(* IEC 61131-3 sources: plcassist-cli/packages/volt-lsp-iec/test-corpus/awa-palletizer/Device/Plc Logic/Application/Library Manager/ElementCollections, 110 files *)

(* ---- CONSTANTS.gvl ---- *)
VAR_GLOBAL
	GC_TREENODEFACTORY : TreeNodeFactory := STRUCT();
	GC_LINKEDOBJECTREFERENCEFACTORY : LinkedObjectReferenceFactory := STRUCT();
END_VAR

(* ---- VARIABLES.gvl ---- *)
VAR_GLOBAL
	G_LOCKWAITTIME : SYSTIME := 300;
	G_NULLELEMENT : NullElement;
END_VAR

(* ---- IBOOLELEMENT.itf ---- *)
INTERFACE IBOOLELEMENT
END_INTERFACE

(* ---- ICOLLECTION.itf ---- *)
INTERFACE ICOLLECTION
END_INTERFACE

METHOD ADDELEMENT : COLLECTION_ERROR
VAR_INPUT
	ITFELEMENT : IElement;
END_VAR
END_METHOD

METHOD CONTAINSELEMENT : COLLECTION_ERROR
VAR_INPUT
	ITFELEMENT : IElement;
END_VAR
VAR_OUTPUT
	XRESULT : BOOL;
END_VAR
END_METHOD

METHOD COUNTELEMENTS : UDINT
END_METHOD

METHOD ELEMENTITERATOR : COLLECTION_ERROR
VAR_INPUT
	ITFITERATOR : IIterator;
END_VAR
END_METHOD

METHOD REMOVEALLELEMENTS : COLLECTION_ERROR
END_METHOD

METHOD REMOVEELEMENT : COLLECTION_ERROR
VAR_INPUT
	ITFELEMENT : IElement;
END_VAR
END_METHOD

(* ---- ICONTAINSVALUE.itf ---- *)
INTERFACE ICONTAINSVALUE
END_INTERFACE

METHOD CONTAINSVALUE : COLLECTION_ERROR
VAR_INPUT
	ITFELEMENT : IElement;
END_VAR
VAR_OUTPUT
	XRESULT : BOOL;
END_VAR
END_METHOD

(* ---- IDINTELEMENT.itf ---- *)
INTERFACE IDINTELEMENT
END_INTERFACE

(* ---- IDOUBLELINKEDLIST.itf ---- *)
INTERFACE IDOUBLELINKEDLIST
END_INTERFACE

METHOD REMOVEFIRSTELEMENT : COLLECTION_ERROR
END_METHOD

METHOD REMOVELASTELEMENT : COLLECTION_ERROR
END_METHOD

(* ---- IDOUBLELINKEDLIST2.itf ---- *)
INTERFACE IDOUBLELINKEDLIST2
END_INTERFACE

METHOD SAFEELEMENTITERATOR : COLLECTION_ERROR
VAR_INPUT
	ITFITERATOR : ISafeLinkedListIterator;
END_VAR
END_METHOD

(* ---- IELEMENT.itf ---- *)
INTERFACE IELEMENT
END_INTERFACE

METHOD ELEMENTCOMPARETO : INT
VAR_INPUT
	ITFELEMENT : IElement;
END_VAR
END_METHOD

METHOD ELEMENTEQUALS : BOOL
VAR_INPUT
	ITFELEMENT : IElement;
END_VAR
END_METHOD

METHOD ELEMENTHASHCODE : LINT
END_METHOD

(* ---- IINTELEMENT.itf ---- *)
INTERFACE IINTELEMENT
END_INTERFACE

(* ---- IITERATOR.itf ---- *)
INTERFACE IITERATOR
END_INTERFACE

METHOD HASNEXT : BOOL
END_METHOD

METHOD NEXT : COLLECTION_ERROR
VAR_OUTPUT
	ITFELEMENT : IElement;
END_VAR
END_METHOD

(* ---- ILINKEDLISTITERATOR.itf ---- *)
INTERFACE ILINKEDLISTITERATOR
END_INTERFACE

(* ---- ILINKEDOBJECTREFERENCE.itf ---- *)
INTERFACE ILINKEDOBJECTREFERENCE
END_INTERFACE

(* ---- ILINTELEMENT.itf ---- *)
INTERFACE ILINTELEMENT
END_INTERFACE

(* ---- ILIST.itf ---- *)
INTERFACE ILIST
END_INTERFACE

METHOD GETELEMENTAT : COLLECTION_ERROR
VAR_INPUT
	UDIPOSITION : UDINT;
END_VAR
VAR_OUTPUT
	ITFELEMENT : IElement;
END_VAR
END_METHOD

METHOD GETELEMENTPOSITION : COLLECTION_ERROR
VAR_INPUT
	ITFELEMENT : IElement;
END_VAR
VAR_OUTPUT
	UDIPOSITION : UDINT;
END_VAR
END_METHOD

METHOD INSERTELEMENTAT : COLLECTION_ERROR
VAR_INPUT
	UDIPOSITION : UDINT;
	ITFELEMENT : IElement;
END_VAR
END_METHOD

METHOD REMOVEELEMENTAT : COLLECTION_ERROR
VAR_INPUT
	UDIPOSITION : UDINT;
END_VAR
END_METHOD

METHOD SETELEMENTAT : COLLECTION_ERROR
VAR_INPUT
	UDIPOSITION : UDINT;
	ITFELEMENT : IElement;
END_VAR
END_METHOD

(* ---- ILIST2.itf ---- *)
INTERFACE ILIST2
END_INTERFACE

(* ---- ILIST3.itf ---- *)
INTERFACE ILIST3
END_INTERFACE

METHOD SAFEELEMENTITERATOR : COLLECTION_ERROR
VAR_INPUT
	ITFITERATOR : ISafeListIterator;
END_VAR
END_METHOD

(* ---- ILISTITERATOR.itf ---- *)
INTERFACE ILISTITERATOR
END_INTERFACE

(* ---- ILOCKABLE.itf ---- *)
INTERFACE ILOCKABLE
END_INTERFACE

METHOD LOCK : BOOL
END_METHOD

METHOD RELEASELOCK
END_METHOD

(* ---- IMAP.itf ---- *)
INTERFACE IMAP
END_INTERFACE

METHOD ADDKEYVALUEPAIR : COLLECTION_ERROR
VAR_INPUT
	ITFKEY : IElement;
	ITFVALUE : IElement;
END_VAR
END_METHOD

METHOD CONTAINSKEY : COLLECTION_ERROR
VAR_INPUT
	ITFKEY : IElement;
END_VAR
VAR_OUTPUT
	XRESULT : BOOL;
END_VAR
END_METHOD

METHOD COUNTKEYS : UDINT
END_METHOD

METHOD GETELEMENTBYKEY : COLLECTION_ERROR
VAR_INPUT
	ITFKEY : IElement;
END_VAR
VAR_OUTPUT
	ITFVALUE : IElement;
END_VAR
END_METHOD

METHOD KEYS : COLLECTION_ERROR
VAR_INPUT
	ITFITERATOR : IIterator;
END_VAR
END_METHOD

METHOD REMOVEBYKEY : COLLECTION_ERROR
VAR_INPUT
	ITFKEY : IElement;
END_VAR
END_METHOD

METHOD VALUES : COLLECTION_ERROR
VAR_INPUT
	ITFITERATOR : IIterator;
END_VAR
END_METHOD

(* ---- IMAP2.itf ---- *)
INTERFACE IMAP2
END_INTERFACE

METHOD REMOVEALLELEMENTS : COLLECTION_ERROR
END_METHOD

(* ---- IMAP3.itf ---- *)
INTERFACE IMAP3
END_INTERFACE

METHOD SAFEKEYS : COLLECTION_ERROR
VAR_INPUT
	ITFITERATOR : ISafeListIterator;
END_VAR
END_METHOD

METHOD SAFEVALUES : COLLECTION_ERROR
VAR_INPUT
	ITFITERATOR : ISafeListIterator;
END_VAR
END_METHOD

(* ---- IMODCOUNTER.itf ---- *)
INTERFACE IMODCOUNTER
END_INTERFACE

(* ---- INULLELEMENT.itf ---- *)
INTERFACE INULLELEMENT
END_INTERFACE

(* ---- IOBJECTREFERENCE.itf ---- *)
INTERFACE IOBJECTREFERENCE
END_INTERFACE

(* ---- IONLINECHANGESAFELINKEDLISTELEMENT.itf ---- *)
INTERFACE IONLINECHANGESAFELINKEDLISTELEMENT
END_INTERFACE

METHOD UPDATEELEMENT
VAR_INPUT
	ITFELEMENT : IElement;
END_VAR
END_METHOD

(* ---- IQUEUE.itf ---- *)
INTERFACE IQUEUE
END_INTERFACE

METHOD PEEK : COLLECTION_ERROR
VAR_OUTPUT
	ITFELEMENT : IElement;
END_VAR
END_METHOD

METHOD POLL : COLLECTION_ERROR
VAR_OUTPUT
	ITFELEMENT : IElement;
END_VAR
END_METHOD

(* ---- IQUEUE2.itf ---- *)
INTERFACE IQUEUE2
END_INTERFACE

(* ---- IQUEUE3.itf ---- *)
INTERFACE IQUEUE3
END_INTERFACE

METHOD SAFEELEMENTITERATOR : COLLECTION_ERROR
VAR_INPUT
	ITFITERATOR : ISafeListIterator;
END_VAR
END_METHOD

(* ---- ISAFEITERATOR.itf ---- *)
INTERFACE ISAFEITERATOR
END_INTERFACE

METHOD NEXT : COLLECTION_ERROR
VAR_OUTPUT
	ITFELEMENT : IElement;
END_VAR
END_METHOD

(* ---- ISAFELINKEDLISTITERATOR.itf ---- *)
INTERFACE ISAFELINKEDLISTITERATOR
END_INTERFACE

(* ---- ISAFELISTITERATOR.itf ---- *)
INTERFACE ISAFELISTITERATOR
END_INTERFACE

(* ---- ISORTEDLIST.itf ---- *)
INTERFACE ISORTEDLIST
END_INTERFACE

METHOD ADDELEMENTWITHOUTSORTING : COLLECTION_ERROR
VAR_INPUT
	ITFELEMENT : IElement;
END_VAR
END_METHOD

METHOD SORT : COLLECTION_ERROR
END_METHOD

(* ---- ISORTEDLIST2.itf ---- *)
INTERFACE ISORTEDLIST2
END_INTERFACE

(* ---- ISORTEDLIST3.itf ---- *)
INTERFACE ISORTEDLIST3
END_INTERFACE

METHOD SAFEELEMENTITERATOR : COLLECTION_ERROR
VAR_INPUT
	ITFITERATOR : ISafeListIterator;
END_VAR
END_METHOD

(* ---- ISTACK.itf ---- *)
INTERFACE ISTACK
END_INTERFACE

METHOD PEEK : COLLECTION_ERROR
VAR_OUTPUT
	ITFELEMENT : IElement;
END_VAR
END_METHOD

METHOD POP : COLLECTION_ERROR
VAR_OUTPUT
	ITFELEMENT : IElement;
END_VAR
END_METHOD

(* ---- ISTACK2.itf ---- *)
INTERFACE ISTACK2
END_INTERFACE

(* ---- ISTACK3.itf ---- *)
INTERFACE ISTACK3
END_INTERFACE

METHOD SAFEELEMENTITERATOR : COLLECTION_ERROR
VAR_INPUT
	ITFITERATOR : ISafeListIterator;
END_VAR
END_METHOD

(* ---- ISTRINGELEMENT.itf ---- *)
INTERFACE ISTRINGELEMENT
END_INTERFACE

(* ---- ITIMEELEMENT.itf ---- *)
INTERFACE ITIMEELEMENT
END_INTERFACE

(* ---- ITREENODE.itf ---- *)
INTERFACE ITREENODE
END_INTERFACE

METHOD ADDCHILD : COLLECTION_ERROR
VAR_INPUT
	ITFELEMENT : IElement;
END_VAR
VAR_OUTPUT
	ITFTREENODE : ITreeNode;
END_VAR
END_METHOD

METHOD CHILDREN : COLLECTION_ERROR
VAR_INPUT
	ITFITERATOR : IIterator;
END_VAR
END_METHOD

METHOD CONTAINSCHILD : COLLECTION_ERROR
VAR_INPUT
	ITFELEMENT : IElement;
END_VAR
VAR_OUTPUT
	XRESULT : BOOL;
END_VAR
END_METHOD

METHOD COUNTCHILDREN : UDINT
END_METHOD

METHOD MOVENODE : COLLECTION_ERROR
VAR_INPUT
	ITFTARGETTREENODE : ITreeNode;
END_VAR
END_METHOD

METHOD PARENT : COLLECTION_ERROR
VAR_OUTPUT
	ITFPARENT : ITreeNode;
END_VAR
END_METHOD

METHOD REMOVECHILD : COLLECTION_ERROR
VAR_INPUT
	ITFELEMENT : IElement;
END_VAR
END_METHOD

METHOD ROOTNODE : COLLECTION_ERROR
VAR_OUTPUT
	ITFROOTNODE : ITreeNode;
END_VAR
END_METHOD

(* ---- ITREENODE2.itf ---- *)
INTERFACE ITREENODE2
END_INTERFACE

METHOD SAFECHILDREN : COLLECTION_ERROR
VAR_INPUT
	ITFITERATOR : ISafeLinkedListIterator;
END_VAR
END_METHOD

(* ---- IUDINTELEMENT.itf ---- *)
INTERFACE IUDINTELEMENT
END_INTERFACE

(* ---- IUINTELEMENT.itf ---- *)
INTERFACE IUINTELEMENT
END_INTERFACE

(* ---- IULINTELEMENT.itf ---- *)
INTERFACE IULINTELEMENT
END_INTERFACE

(* ---- IWSTRINGELEMENT.itf ---- *)
INTERFACE IWSTRINGELEMENT
END_INTERFACE

(* ---- COMPARESTRING.fun ---- *)
FUNCTION COMPARESTRING : INT
VAR_INPUT
	PS1 : POINTER TO STRING;
	PS2 : POINTER TO STRING;
END_VAR
END_FUNCTION

(* ---- COMPAREWSTRING.fun ---- *)
FUNCTION COMPAREWSTRING : INT
VAR_INPUT
	PW1 : POINTER TO WSTRING;
	PW2 : POINTER TO WSTRING;
END_VAR
END_FUNCTION

(* ---- GETLIBVERSION.fun ---- *)
FUNCTION GETLIBVERSION : VERSION
END_FUNCTION

(* ---- GETLIBVERSIONNUMBER.fun ---- *)
FUNCTION GETLIBVERSIONNUMBER : DWORD
END_FUNCTION

(* ---- HASHCODEFROMSTRING.fun ---- *)
FUNCTION HASHCODEFROMSTRING : UDINT
VAR_INPUT
	PSIN : POINTER TO STRING;
END_VAR
END_FUNCTION

(* ---- HASHCODEFROMWSTRING.fun ---- *)
FUNCTION HASHCODEFROMWSTRING : UDINT
VAR_INPUT
	PWIN : POINTER TO WSTRING;
END_VAR
END_FUNCTION

(* ---- ISLIBRELEASED.fun ---- *)
FUNCTION ISLIBRELEASED : BOOL
END_FUNCTION

(* ---- BOOLDATA.fb ---- *)
FUNCTION_BLOCK BOOLDATA EXTENDS InstanceData
VAR_INPUT
	XVALUE : BOOL;
END_VAR
END_FUNCTION_BLOCK

(* ---- BOOLELEMENT.fb ---- *)
FUNCTION_BLOCK BOOLELEMENT EXTENDS InstanceBase
VAR_INPUT
	XVALUE : BOOL;
END_VAR
VAR
	BOOLVALUE : BOOL;
END_VAR
END_FUNCTION_BLOCK

METHOD ELEMENTCOMPARETO : INT
VAR_INPUT
	ITFELEMENT : IElement;
END_VAR
END_METHOD

METHOD ELEMENTEQUALS : BOOL
VAR_INPUT
	ITFELEMENT : IElement;
END_VAR
END_METHOD

METHOD ELEMENTHASHCODE : LINT
END_METHOD

METHOD PRVINSTINIT : FBF.ERROR
VAR_INPUT
	ITFDATA : FBF.IData;
END_VAR
END_METHOD

(* ---- BOOLELEMENTFACTORY.fb ---- *)
FUNCTION_BLOCK BOOLELEMENTFACTORY EXTENDS FactoryBase
VAR
	PRVINSTCOUNT : CAA.COUNT;
	PRVINSTPOOLEXTENDSFACTOR : USINT;
	PRVINSTSIZE : CAA.SIZE;
END_VAR
END_FUNCTION_BLOCK

METHOD CREATE : IBoolElement
VAR_INPUT
	XVALUE : BOOL;
END_VAR
VAR_OUTPUT
	EERROR : FBF.ERROR;
END_VAR
END_METHOD

(* ---- DINTDATA.fb ---- *)
FUNCTION_BLOCK DINTDATA EXTENDS InstanceData
VAR_INPUT
	DIVALUE : DINT;
END_VAR
END_FUNCTION_BLOCK

(* ---- DINTELEMENT.fb ---- *)
FUNCTION_BLOCK DINTELEMENT EXTENDS InstanceBase
VAR_INPUT
	DIVALUE : DINT;
END_VAR
VAR
	DINTVALUE : DINT;
END_VAR
END_FUNCTION_BLOCK

METHOD ELEMENTCOMPARETO : INT
VAR_INPUT
	ITFELEMENT : IElement;
END_VAR
END_METHOD

METHOD ELEMENTEQUALS : BOOL
VAR_INPUT
	ITFELEMENT : IElement;
END_VAR
END_METHOD

METHOD ELEMENTHASHCODE : LINT
END_METHOD

METHOD PRVINSTINIT : FBF.ERROR
VAR_INPUT
	ITFDATA : FBF.IData;
END_VAR
END_METHOD

(* ---- DINTELEMENTFACTORY.fb ---- *)
FUNCTION_BLOCK DINTELEMENTFACTORY EXTENDS FactoryBase
VAR
	PRVINSTCOUNT : CAA.COUNT;
	PRVINSTPOOLEXTENDSFACTOR : USINT;
	PRVINSTSIZE : CAA.SIZE;
END_VAR
END_FUNCTION_BLOCK

METHOD CREATE : IDintElement
VAR_INPUT
	DIVALUE : DINT;
END_VAR
VAR_OUTPUT
	EERROR : FBF.ERROR;
END_VAR
END_METHOD

(* ---- HASHTABLE.fb ---- *)
FUNCTION_BLOCK HASHTABLE EXTENDS InstanceBase
VAR_INPUT
	PAELEMENTS : POINTER TO KeyValuePair;
	PALINKEDELEMENTS : POINTER TO KeyValuePair;
	PAITERATORELEMENTS : POINTER TO IElement;
	UDIMAXELEMENTS : UDINT;
END_VAR
VAR
	_UDICOUNT : UDINT;
	_XWPOINTERTOTHIS : __XWORD := THIS;
	_BYLOCK : BYTE;
	_ULINTCOUNTMODS : ULINT;
	_UIGROWFACTOR : UINT := 1;
	_UIPREALLOCATION : UINT := 100;
	_LOCKWAITTIME : SYSTIME := Variables.g_LockWaitTime;
	COUNTMODIFICATIONS : ULINT;
	LOCKWAITTIME : SYSTIME;
END_VAR
END_FUNCTION_BLOCK

METHOD ADDKEYVALUEPAIR : COLLECTION_ERROR
VAR_INPUT
	ITFKEY : IElement;
	ITFVALUE : IElement;
END_VAR
END_METHOD

METHOD ADDKEYVALUEPAIRINTERNAL : COLLECTION_ERROR
VAR_INPUT
	ITFKEY : IElement;
	ITFVALUE : IElement;
	XINCREF : BOOL;
END_VAR
END_METHOD

METHOD CONTAINSKEY : COLLECTION_ERROR
VAR_INPUT
	ITFKEY : IElement;
END_VAR
VAR_OUTPUT
	XRESULT : BOOL;
END_VAR
END_METHOD

METHOD CONTAINSKEYINTERNAL : COLLECTION_ERROR
VAR_INPUT
	ITFKEY : IElement;
END_VAR
VAR_OUTPUT
	XRESULT : BOOL;
END_VAR
END_METHOD

METHOD COUNTKEYS : UDINT
END_METHOD

METHOD DISPOSE : BOOL
END_METHOD

METHOD ELEMENTCOMPARETO : INT
VAR_INPUT
	ITFELEMENT : IElement;
END_VAR
END_METHOD

METHOD ELEMENTEQUALS : BOOL
VAR_INPUT
	ITFELEMENT : IElement;
END_VAR
END_METHOD

METHOD ELEMENTHASHCODE : LINT
END_METHOD

METHOD GETARRAYINDEX : UDINT
VAR_INPUT
	ITFKEY : IElement;
END_VAR
END_METHOD

METHOD GETELEMENTBYKEY : COLLECTION_ERROR
VAR_INPUT
	ITFKEY : IElement;
END_VAR
VAR_OUTPUT
	ITFVALUE : IElement;
END_VAR
END_METHOD

METHOD KEYS : COLLECTION_ERROR
VAR_INPUT
	ITFITERATOR : IIterator;
END_VAR
END_METHOD

METHOD LOCK : BOOL
END_METHOD

METHOD NEXTFREELINKEDELEMENT : COLLECTION_ERROR
VAR_OUTPUT
	PKEYVALUEPAIR : POINTER TO KeyValuePair;
END_VAR
END_METHOD

METHOD REALLOC : BOOL
END_METHOD

METHOD RELEASELOCK
END_METHOD

METHOD REMOVEALLELEMENTS : COLLECTION_ERROR
END_METHOD

METHOD REMOVEBYKEY : COLLECTION_ERROR
VAR_INPUT
	ITFKEY : IElement;
END_VAR
END_METHOD

METHOD SAFEKEYS : COLLECTION_ERROR
VAR_INPUT
	ITFITERATOR : ISafeListIterator;
END_VAR
END_METHOD

METHOD SAFEVALUES : COLLECTION_ERROR
VAR_INPUT
	ITFITERATOR : ISafeListIterator;
END_VAR
END_METHOD

METHOD VALUES : COLLECTION_ERROR
VAR_INPUT
	ITFITERATOR : IIterator;
END_VAR
END_METHOD

METHOD PRVINSTINIT : FBF.ERROR
VAR_INPUT
	ITFDATA : FBF.IData;
END_VAR
END_METHOD

(* ---- HASHTABLEARGS.fb ---- *)
FUNCTION_BLOCK HASHTABLEARGS EXTENDS InstanceData
VAR_INPUT
	PAELEMENTS : POINTER TO KeyValuePair;
	PALINKEDELEMENTS : POINTER TO KeyValuePair;
	PAITERATORELEMENTS : POINTER TO IElement;
	UDIMAXELEMENTS : UDINT;
	UIGROWFACTOR : UINT;
	UIPREALLOCATION : UINT;
END_VAR
END_FUNCTION_BLOCK

(* ---- HASHTABLEFACTORY.fb ---- *)
FUNCTION_BLOCK HASHTABLEFACTORY EXTENDS FactoryBase
VAR
	PRVINSTCOUNT : CAA.COUNT;
	PRVINSTPOOLEXTENDSFACTOR : USINT;
	PRVINSTSIZE : CAA.SIZE;
END_VAR
END_FUNCTION_BLOCK

METHOD CREATE : IMap3
VAR_INPUT
	UDIMAXELEMENTS : UDINT;
END_VAR
VAR_OUTPUT
	EERROR : FBF.ERROR;
END_VAR
END_METHOD

METHOD CREATEDYNAMICHASHTABLE : IMap2
VAR_INPUT
	UDIINITIALSIZE : UDINT;
	UIGROWFACTOR : UINT;
END_VAR
VAR_OUTPUT
	EERROR : FBF.ERROR;
END_VAR
END_METHOD

METHOD CREATEDYNAMICHASHTABLEPREALLOC : IMap2
VAR_INPUT
	UDIINITIALSIZE : UDINT;
	UIGROWFACTOR : UINT;
	UIPREALLOCATION : UINT;
END_VAR
VAR_OUTPUT
	EERROR : FBF.ERROR;
END_VAR
END_METHOD

(* ---- INTDATA.fb ---- *)
FUNCTION_BLOCK INTDATA EXTENDS InstanceData
VAR_INPUT
	IVALUE : INT;
END_VAR
END_FUNCTION_BLOCK

(* ---- INTELEMENT.fb ---- *)
FUNCTION_BLOCK INTELEMENT EXTENDS InstanceBase
VAR_INPUT
	IVALUE : INT;
END_VAR
VAR
	INTVALUE : INT;
END_VAR
END_FUNCTION_BLOCK

METHOD ELEMENTCOMPARETO : INT
VAR_INPUT
	ITFELEMENT : IElement;
END_VAR
END_METHOD

METHOD ELEMENTEQUALS : BOOL
VAR_INPUT
	ITFELEMENT : IElement;
END_VAR
END_METHOD

METHOD ELEMENTHASHCODE : LINT
END_METHOD

METHOD PRVINSTINIT : FBF.ERROR
VAR_INPUT
	ITFDATA : FBF.IData;
END_VAR
END_METHOD

(* ---- INTELEMENTFACTORY.fb ---- *)
FUNCTION_BLOCK INTELEMENTFACTORY EXTENDS FactoryBase
VAR
	PRVINSTCOUNT : CAA.COUNT;
	PRVINSTPOOLEXTENDSFACTOR : USINT;
	PRVINSTSIZE : CAA.SIZE;
END_VAR
END_FUNCTION_BLOCK

METHOD CREATE : IIntElement
VAR_INPUT
	IVALUE : INT;
END_VAR
VAR_OUTPUT
	EERROR : FBF.ERROR;
END_VAR
END_METHOD

(* ---- LINKEDLIST.fb ---- *)
FUNCTION_BLOCK LINKEDLIST EXTENDS InstanceBase
VAR
	_SNAME : STRING := 'LinkedList';
	_RESULT : RTS_IEC_RESULT;
	_XWPOINTERTOTHIS : __XWORD := THIS;
	_BYLOCK : BYTE;
	_ULINTCOUNTMODS : ULINT;
	_ITFFIRSTLINKEDOBJECTREFERENCE : ILinkedObjectReference := 0;
	_ITFLASTLINKEDOBJECTREFERENCE : ILinkedObjectReference := 0;
	_UDICOUNT : UDINT;
	_LOCKWAITTIME : SYSTIME := Variables.g_LockWaitTime;
	COUNTMODIFICATIONS : ULINT;
	LOCKWAITTIME : SYSTIME;
END_VAR
END_FUNCTION_BLOCK

METHOD ADDELEMENT : COLLECTION_ERROR
VAR_INPUT
	ITFELEMENT : IElement;
END_VAR
END_METHOD

METHOD ADDELEMENTINTERNAL : COLLECTION_ERROR
VAR_INPUT
	ITFELEMENT : IElement;
	XINCREMENTREFERENCECOUNTER : BOOL;
END_VAR
END_METHOD

METHOD CONTAINSELEMENT : COLLECTION_ERROR
VAR_INPUT
	ITFELEMENT : IElement;
END_VAR
VAR_OUTPUT
	XRESULT : BOOL;
END_VAR
END_METHOD

METHOD COUNTELEMENTS : UDINT
END_METHOD

METHOD DISPOSE : BOOL
END_METHOD

METHOD ELEMENTCOMPARETO : INT
VAR_INPUT
	ITFELEMENT : IElement;
END_VAR
END_METHOD

METHOD ELEMENTEQUALS : BOOL
VAR_INPUT
	ITFELEMENT : IElement;
END_VAR
END_METHOD

METHOD ELEMENTHASHCODE : LINT
END_METHOD

METHOD ELEMENTITERATOR : COLLECTION_ERROR
VAR_INPUT
	ITFITERATOR : IIterator;
END_VAR
END_METHOD

METHOD LOCK : BOOL
END_METHOD

METHOD RELEASELOCK
END_METHOD

METHOD REMOVEALLELEMENTS : COLLECTION_ERROR
END_METHOD

METHOD REMOVEELEMENT : COLLECTION_ERROR
VAR_INPUT
	ITFELEMENT : IElement;
END_VAR
END_METHOD

METHOD REMOVEELEMENTINTERNAL : COLLECTION_ERROR
VAR_INPUT
	ITFELEMENT : IElement;
	XDECREMENTREFERENCECOUNTER : BOOL;
END_VAR
END_METHOD

METHOD REMOVEFIRSTELEMENT : COLLECTION_ERROR
END_METHOD

METHOD REMOVELASTELEMENT : COLLECTION_ERROR
END_METHOD

METHOD SAFEELEMENTITERATOR : COLLECTION_ERROR
VAR_INPUT
	ITFITERATOR : ISafeLinkedListIterator;
END_VAR
END_METHOD

METHOD PRVINSTINIT : FBF.ERROR
VAR_INPUT
	ITFDATA : FBF.IData;
END_VAR
END_METHOD

(* ---- LINKEDLISTARGS.fb ---- *)
FUNCTION_BLOCK LINKEDLISTARGS EXTENDS InstanceData
END_FUNCTION_BLOCK

(* ---- LINKEDLISTELEMENTBASE.fb ---- *)
FUNCTION_BLOCK LINKEDLISTELEMENTBASE EXTENDS InstanceBase
VAR
	_ITFOBJECTREFERENCE : IObjectReference;
	OBJECTREFERENCE : IObjectReference;
END_VAR
END_FUNCTION_BLOCK

METHOD ELEMENTCOMPARETO : INT
VAR_INPUT
	ITFELEMENT : IElement;
END_VAR
END_METHOD

METHOD ELEMENTEQUALS : BOOL
VAR_INPUT
	ITFELEMENT : IElement;
END_VAR
END_METHOD

METHOD ELEMENTHASHCODE : LINT
END_METHOD

METHOD UPDATEELEMENT
VAR_INPUT
	ITFELEMENT : IElement;
END_VAR
END_METHOD

(* ---- LINKEDLISTFACTORY.fb ---- *)
FUNCTION_BLOCK LINKEDLISTFACTORY EXTENDS FactoryBase
VAR
	PRVINSTCOUNT : CAA.COUNT;
	PRVINSTPOOLEXTENDSFACTOR : USINT;
	PRVINSTSIZE : CAA.SIZE;
END_VAR
END_FUNCTION_BLOCK

METHOD CREATE : IDoubleLinkedList2
VAR_OUTPUT
	EERROR : FBF.ERROR;
END_VAR
END_METHOD

(* ---- LINKEDLISTITERATOR.fb ---- *)
FUNCTION_BLOCK LINKEDLISTITERATOR
VAR
	_ITFLINKEDLISTITERATOR : ILinkedObjectReference;
	_MODCOUNTER : IModCounter;
	_ULINTSTARTMODCOUNT : ULINT;
	_XINVALIDDATA : BOOL;
	FIRSTOBJECTREFERENCE : ILinkedObjectReference;
	MODCOUNTER : IModCounter;
END_VAR
END_FUNCTION_BLOCK

METHOD HASNEXT : BOOL
END_METHOD

METHOD NEXT : COLLECTION_ERROR
VAR_OUTPUT
	ITFELEMENT : IElement;
END_VAR
END_METHOD

(* ---- LINKEDOBJECTREFERENCE.fb ---- *)
FUNCTION_BLOCK LINKEDOBJECTREFERENCE EXTENDS InstanceBase
VAR
	_ITFELEMENT : IElement;
	_ITFLASTLINKEDOBJECTREFERENCE : ILinkedObjectReference;
	_ITFNEXTLINKEDOBJECTREFERENCE : ILinkedObjectReference;
	ELEMENT : IElement;
	LAST : ILinkedObjectReference;
	NEXT : ILinkedObjectReference;
END_VAR
END_FUNCTION_BLOCK

METHOD PRVINSTINIT : FBF.ERROR
VAR_INPUT
	ITFDATA : FBF.IData;
END_VAR
END_METHOD

(* ---- LINKEDOBJECTREFERENCEARGS.fb ---- *)
FUNCTION_BLOCK LINKEDOBJECTREFERENCEARGS EXTENDS InstanceData
END_FUNCTION_BLOCK

(* ---- LINKEDOBJECTREFERENCEFACTORY.fb ---- *)
FUNCTION_BLOCK LINKEDOBJECTREFERENCEFACTORY EXTENDS FactoryBase
VAR
	PRVINSTCOUNT : CAA.COUNT;
	PRVINSTPOOLEXTENDSFACTOR : USINT;
	PRVINSTSIZE : CAA.SIZE;
END_VAR
END_FUNCTION_BLOCK

METHOD CREATE : ILinkedObjectReference
VAR_OUTPUT
	EERROR : FBF.ERROR;
END_VAR
END_METHOD

(* ---- LINTDATA.fb ---- *)
FUNCTION_BLOCK LINTDATA EXTENDS InstanceData
VAR_INPUT
	LIVALUE : LINT;
END_VAR
END_FUNCTION_BLOCK

(* ---- LINTELEMENT.fb ---- *)
FUNCTION_BLOCK LINTELEMENT EXTENDS InstanceBase
VAR_INPUT
	LIVALUE : LINT;
END_VAR
VAR
	LINTVALUE : LINT;
END_VAR
END_FUNCTION_BLOCK

METHOD ELEMENTCOMPARETO : INT
VAR_INPUT
	ITFELEMENT : IElement;
END_VAR
END_METHOD

METHOD ELEMENTEQUALS : BOOL
VAR_INPUT
	ITFELEMENT : IElement;
END_VAR
END_METHOD

METHOD ELEMENTHASHCODE : LINT
END_METHOD

METHOD PRVINSTINIT : FBF.ERROR
VAR_INPUT
	ITFDATA : FBF.IData;
END_VAR
END_METHOD

(* ---- LINTELEMENTFACTORY.fb ---- *)
FUNCTION_BLOCK LINTELEMENTFACTORY EXTENDS FactoryBase
VAR
	PRVINSTCOUNT : CAA.COUNT;
	PRVINSTPOOLEXTENDSFACTOR : USINT;
	PRVINSTSIZE : CAA.SIZE;
END_VAR
END_FUNCTION_BLOCK

METHOD CREATE : ILintElement
VAR_INPUT
	LIVALUE : LINT;
END_VAR
VAR_OUTPUT
	EERROR : FBF.ERROR;
END_VAR
END_METHOD

(* ---- LIST.fb ---- *)
FUNCTION_BLOCK LIST EXTENDS InstanceBase
VAR_INPUT
	PAELEMENTS : POINTER TO IElement;
	UDIMAXELEMENTS : UDINT;
END_VAR
VAR
	_DIMAXPOSITION : DINT := -1;
	_SNAME : STRING := 'List';
	RESULT : RTS_IEC_RESULT;
	_XWPOINTERTOTHIS : __XWORD := THIS;
	_BYLOCK : BYTE;
	_ULINTCOUNTMODS : ULINT;
	_UIGROWFACTOR : UINT := 1;
	_LOCKWAITTIME : SYSTIME := Variables.g_LockWaitTime;
	COUNTMODIFICATIONS : ULINT;
	LOCKWAITTIME : SYSTIME;
END_VAR
END_FUNCTION_BLOCK

METHOD ADDELEMENT : COLLECTION_ERROR
VAR_INPUT
	ITFELEMENT : IElement;
END_VAR
END_METHOD

METHOD CONTAINSELEMENT : COLLECTION_ERROR
VAR_INPUT
	ITFELEMENT : IElement;
END_VAR
VAR_OUTPUT
	XRESULT : BOOL;
END_VAR
END_METHOD

METHOD CONTAINSVALUE : COLLECTION_ERROR
VAR_INPUT
	ITFELEMENT : IElement;
END_VAR
VAR_OUTPUT
	XRESULT : BOOL;
END_VAR
END_METHOD

METHOD COUNTELEMENTS : UDINT
END_METHOD

METHOD DISPOSE : BOOL
END_METHOD

METHOD ELEMENTCOMPARETO : INT
VAR_INPUT
	ITFELEMENT : IElement;
END_VAR
END_METHOD

METHOD ELEMENTEQUALS : BOOL
VAR_INPUT
	ITFELEMENT : IElement;
END_VAR
END_METHOD

METHOD ELEMENTHASHCODE : LINT
END_METHOD

METHOD ELEMENTITERATOR : COLLECTION_ERROR
VAR_INPUT
	ITFITERATOR : IIterator;
END_VAR
END_METHOD

METHOD GETELEMENTAT : COLLECTION_ERROR
VAR_INPUT
	UDIPOSITION : UDINT;
END_VAR
VAR_OUTPUT
	ITFELEMENT : IElement;
END_VAR
END_METHOD

METHOD GETELEMENTPOSITION : COLLECTION_ERROR
VAR_INPUT
	ITFELEMENT : IElement;
END_VAR
VAR_OUTPUT
	UDIPOSITION : UDINT;
END_VAR
END_METHOD

METHOD INSERTELEMENTAT : COLLECTION_ERROR
VAR_INPUT
	UDIPOSITION : UDINT;
	ITFELEMENT : IElement;
END_VAR
END_METHOD

METHOD LOCK : BOOL
END_METHOD

METHOD REALLOC : BOOL
END_METHOD

METHOD RELEASELOCK
END_METHOD

METHOD REMOVEALLELEMENTS : COLLECTION_ERROR
END_METHOD

METHOD REMOVEALLELEMENTSINTERNAL : COLLECTION_ERROR
END_METHOD

METHOD REMOVEELEMENT : COLLECTION_ERROR
VAR_INPUT
	ITFELEMENT : IElement;
END_VAR
END_METHOD

METHOD REMOVEELEMENTAT : COLLECTION_ERROR
VAR_INPUT
	UDIPOSITION : UDINT;
END_VAR
END_METHOD

METHOD REMOVEELEMENTATINTERNAL : COLLECTION_ERROR
VAR_INPUT
	UDIPOSITION : UDINT;
END_VAR
END_METHOD

METHOD SAFEELEMENTITERATOR : COLLECTION_ERROR
VAR_INPUT
	ITFITERATOR : ISafeListIterator;
END_VAR
END_METHOD

METHOD SETELEMENTAT : COLLECTION_ERROR
VAR_INPUT
	UDIPOSITION : UDINT;
	ITFELEMENT : IElement;
END_VAR
END_METHOD

METHOD PRVINSTINIT : FBF.ERROR
VAR_INPUT
	ITFDATA : FBF.IData;
END_VAR
END_METHOD

(* ---- LISTARGS.fb ---- *)
FUNCTION_BLOCK LISTARGS EXTENDS InstanceData
VAR_INPUT
	PAELEMENTS : POINTER TO IElement;
	UDIMAXELEMENTS : UDINT;
	UIGROWFACTOR : UINT;
END_VAR
END_FUNCTION_BLOCK

(* ---- LISTFACTORY.fb ---- *)
FUNCTION_BLOCK LISTFACTORY EXTENDS FactoryBase
VAR
	PRVINSTCOUNT : CAA.COUNT;
	PRVINSTPOOLEXTENDSFACTOR : USINT;
	PRVINSTSIZE : CAA.SIZE;
END_VAR
END_FUNCTION_BLOCK

METHOD CREATE : IList3
VAR_INPUT
	UDIMAXELEMENTS : UDINT;
END_VAR
VAR_OUTPUT
	EERROR : FBF.ERROR;
END_VAR
END_METHOD

METHOD CREATEDYNAMICLIST : IList2
VAR_INPUT
	UDIINITIALSIZE : UDINT;
	UIGROWFACTOR : UINT;
END_VAR
VAR_OUTPUT
	EERROR : FBF.ERROR;
END_VAR
END_METHOD

(* ---- LISTITERATOR.fb ---- *)
FUNCTION_BLOCK LISTITERATOR
VAR
	_DICOUNT : DINT := -1;
	_PAELEMENTS : POINTER TO IElement := 0;
	_DISIZE : DINT;
	_MODCOUNTER : IModCounter;
	_ULINTSTARTMODCOUNT : ULINT;
	ELEMENTARRAY : POINTER TO IElement;
	ELEMENTARRAYSIZE : DINT;
	MODCOUNTER : IModCounter;
END_VAR
END_FUNCTION_BLOCK

METHOD HASNEXT : BOOL
END_METHOD

METHOD NEXT : COLLECTION_ERROR
VAR_OUTPUT
	ITFELEMENT : IElement;
END_VAR
END_METHOD

(* ---- NULLELEMENT.fb ---- *)
FUNCTION_BLOCK NULLELEMENT
END_FUNCTION_BLOCK

METHOD ELEMENTCOMPARETO : INT
VAR_INPUT
	ITFELEMENT : IElement;
END_VAR
END_METHOD

METHOD ELEMENTEQUALS : BOOL
VAR_INPUT
	ITFELEMENT : IElement;
END_VAR
END_METHOD

METHOD ELEMENTHASHCODE : LINT
END_METHOD

(* ---- QUEUE.fb ---- *)
FUNCTION_BLOCK QUEUE EXTENDS InstanceBase
VAR_INPUT
	PAELEMENTS : POINTER TO IElement;
	UDIMAXELEMENTS : UDINT;
END_VAR
VAR
	_DIMAXREARPOSITION : DINT := -1;
	_DIMAXFRONTPOSITION : DINT := -1;
	_SNAME : STRING := 'List';
	RESULT : RTS_IEC_RESULT;
	_XWPOINTERTOTHIS : __XWORD := THIS;
	_BYLOCK : BYTE;
	_ULINTCOUNTMODS : ULINT;
	_UIGROWFACTOR : UINT := 1;
	_LOCKWAITTIME : SYSTIME := Variables.g_LockWaitTime;
	COUNTMODIFICATIONS : ULINT;
	LOCKWAITTIME : SYSTIME;
END_VAR
END_FUNCTION_BLOCK

METHOD ADDELEMENT : COLLECTION_ERROR
VAR_INPUT
	ITFELEMENT : IElement;
END_VAR
END_METHOD

METHOD CONTAINSELEMENT : COLLECTION_ERROR
VAR_INPUT
	ITFELEMENT : IElement;
END_VAR
VAR_OUTPUT
	XRESULT : BOOL;
END_VAR
END_METHOD

METHOD CONTAINSVALUE : COLLECTION_ERROR
VAR_INPUT
	ITFELEMENT : IElement;
END_VAR
VAR_OUTPUT
	XRESULT : BOOL;
END_VAR
END_METHOD

METHOD COUNTELEMENTS : UDINT
END_METHOD

METHOD DISPOSE : BOOL
END_METHOD

METHOD ELEMENTCOMPARETO : INT
VAR_INPUT
	ITFELEMENT : IElement;
END_VAR
END_METHOD

METHOD ELEMENTEQUALS : BOOL
VAR_INPUT
	ITFELEMENT : IElement;
END_VAR
END_METHOD

METHOD ELEMENTHASHCODE : LINT
END_METHOD

METHOD ELEMENTITERATOR : COLLECTION_ERROR
VAR_INPUT
	ITFITERATOR : IIterator;
END_VAR
END_METHOD

METHOD LOCK : BOOL
END_METHOD

METHOD PEEK : COLLECTION_ERROR
VAR_OUTPUT
	ITFELEMENT : IElement;
END_VAR
END_METHOD

METHOD POLL : COLLECTION_ERROR
VAR_OUTPUT
	ITFELEMENT : IElement;
END_VAR
END_METHOD

METHOD REALLOC : BOOL
END_METHOD

METHOD RELEASELOCK
END_METHOD

METHOD REMOVEALLELEMENTS : COLLECTION_ERROR
END_METHOD

METHOD REMOVEALLELEMENTSINTERNAL : COLLECTION_ERROR
END_METHOD

METHOD REMOVEELEMENT : COLLECTION_ERROR
VAR_INPUT
	ITFELEMENT : IElement;
END_VAR
END_METHOD

METHOD REMOVEELEMENTATINTERNAL : COLLECTION_ERROR
VAR_INPUT
	UDIPOSITION : UDINT;
END_VAR
END_METHOD

METHOD SAFEELEMENTITERATOR : COLLECTION_ERROR
VAR_INPUT
	ITFITERATOR : ISafeListIterator;
END_VAR
END_METHOD

METHOD PRVINSTINIT : FBF.ERROR
VAR_INPUT
	ITFDATA : FBF.IData;
END_VAR
END_METHOD

(* ---- QUEUEFACTORY.fb ---- *)
FUNCTION_BLOCK QUEUEFACTORY EXTENDS FactoryBase
VAR
	PRVINSTCOUNT : CAA.COUNT;
	PRVINSTPOOLEXTENDSFACTOR : USINT;
	PRVINSTSIZE : CAA.SIZE;
END_VAR
END_FUNCTION_BLOCK

METHOD CREATE : IQueue3
VAR_INPUT
	UDIMAXELEMENTS : UDINT;
END_VAR
VAR_OUTPUT
	EERROR : FBF.ERROR;
END_VAR
END_METHOD

METHOD CREATEDYNAMICQUEUE : IQueue2
VAR_INPUT
	UDIINITIALSIZE : UDINT;
	UIGROWFACTOR : UINT;
END_VAR
VAR_OUTPUT
	EERROR : FBF.ERROR;
END_VAR
END_METHOD

(* ---- SAFELINKEDLISTITERATOR.fb ---- *)
FUNCTION_BLOCK SAFELINKEDLISTITERATOR
VAR
	_ITFLINKEDLISTITERATOR : ILinkedObjectReference;
	_ITFLASTLINKEDLISTITERATOR : ILinkedObjectReference;
	_MODCOUNTER : IModCounter;
	_ULINTSTARTMODCOUNT : ULINT;
	_XINVALIDDATA : BOOL;
	_ITFLOCKER : ILockable;
	FIRSTOBJECTREFERENCE : ILinkedObjectReference;
	LOCKABLECOLLECTION : ILockable;
	MODCOUNTER : IModCounter;
END_VAR
END_FUNCTION_BLOCK

METHOD NEXT : COLLECTION_ERROR
VAR_OUTPUT
	ITFELEMENT : IElement;
END_VAR
END_METHOD

(* ---- SAFELISTITERATOR.fb ---- *)
FUNCTION_BLOCK SAFELISTITERATOR
VAR
	_DICOUNT : DINT := -1;
	_PAELEMENTS : POINTER TO IElement := 0;
	_DISIZE : DINT;
	_MODCOUNTER : IModCounter;
	_ULINTSTARTMODCOUNT : ULINT;
	_ITFLOCKER : ILockable;
	_ITFLASTELEMENT : IElement := 0;
	ELEMENTARRAY : POINTER TO IElement;
	ELEMENTARRAYSIZE : DINT;
	LOCKABLECOLLECTION : ILockable;
	MODCOUNTER : IModCounter;
END_VAR
END_FUNCTION_BLOCK

METHOD NEXT : COLLECTION_ERROR
VAR_OUTPUT
	ITFELEMENT : IElement;
END_VAR
END_METHOD

(* ---- SORTEDLIST.fb ---- *)
FUNCTION_BLOCK SORTEDLIST EXTENDS InstanceBase
VAR_INPUT
	PAELEMENTS : POINTER TO IElement;
	UDIMAXELEMENTS : UDINT;
	XSORTAFTERONLINECHANGE : BOOL := FALSE;
END_VAR
VAR
	_DIMAXPOSITION : DINT := -1;
	_SNAME : STRING := 'List';
	RESULT : RTS_IEC_RESULT;
	_XWPOINTERTOTHIS : __XWORD := THIS;
	_BYLOCK : BYTE;
	_HEVT_ONLINECHANGEDONE : RTS_IEC_HANDLE;
	_HINTERFACEEVT_ONLINECHANGEDONE : RTS_IEC_HANDLE;
	_ITFEVENTCALLBACK : CmpEventMgr_Interfaces.ICmpEventCallback;
	_ULINTCOUNTMODS : ULINT;
	_UIGROWFACTOR : UINT := 1;
	_LOCKWAITTIME : SYSTIME := Variables.g_LockWaitTime;
	COUNTMODIFICATIONS : ULINT;
	LOCKWAITTIME : SYSTIME;
END_VAR
END_FUNCTION_BLOCK

METHOD ADDELEMENT : COLLECTION_ERROR
VAR_INPUT
	ITFELEMENT : IElement;
END_VAR
END_METHOD

METHOD ADDELEMENTWITHOUTSORTING : COLLECTION_ERROR
VAR_INPUT
	ITFELEMENT : IElement;
END_VAR
END_METHOD

METHOD CONTAINSELEMENT : COLLECTION_ERROR
VAR_INPUT
	ITFELEMENT : IElement;
END_VAR
VAR_OUTPUT
	XRESULT : BOOL;
END_VAR
END_METHOD

METHOD CONTAINSVALUE : COLLECTION_ERROR
VAR_INPUT
	ITFELEMENT : IElement;
END_VAR
VAR_OUTPUT
	XRESULT : BOOL;
END_VAR
END_METHOD

METHOD COUNTELEMENTS : UDINT
END_METHOD

METHOD DISPOSE : BOOL
END_METHOD

METHOD ELEMENTCOMPARETO : INT
VAR_INPUT
	ITFELEMENT : IElement;
END_VAR
END_METHOD

METHOD ELEMENTEQUALS : BOOL
VAR_INPUT
	ITFELEMENT : IElement;
END_VAR
END_METHOD

METHOD ELEMENTHASHCODE : LINT
END_METHOD

METHOD ELEMENTITERATOR : COLLECTION_ERROR
VAR_INPUT
	ITFITERATOR : IIterator;
END_VAR
END_METHOD

METHOD EVENTCALLBACK : UDINT
VAR_INPUT
	PEVENTPARAM : POINTER TO EventParam;
END_VAR
END_METHOD

METHOD FB_INIT : BOOL
VAR_INPUT
	BINITRETAINS : BOOL;
	BINCOPYCODE : BOOL;
END_VAR
END_METHOD

METHOD FB_EXIT : BOOL
VAR_INPUT
	BINCOPYCODE : BOOL;
END_VAR
END_METHOD

METHOD GETELEMENTAT : COLLECTION_ERROR
VAR_INPUT
	UDIPOSITION : UDINT;
END_VAR
VAR_OUTPUT
	ITFELEMENT : IElement;
END_VAR
END_METHOD

METHOD GETELEMENTPOSITION : COLLECTION_ERROR
VAR_INPUT
	ITFELEMENT : IElement;
END_VAR
VAR_OUTPUT
	UDIPOSITION : UDINT;
END_VAR
END_METHOD

METHOD INSERTELEMENTAT : COLLECTION_ERROR
VAR_INPUT
	UDIPOSITION : UDINT;
	ITFELEMENT : IElement;
END_VAR
END_METHOD

METHOD LOCK : BOOL
END_METHOD

METHOD QSORTHELPER : BOOL
VAR_INPUT
	DILEFT : DINT;
	DIRIGHT : DINT;
END_VAR
END_METHOD

METHOD QUICKSORT : BOOL
VAR_INPUT
	DILEFT : DINT;
	DIRIGHT : DINT;
END_VAR
END_METHOD

METHOD REALLOC : BOOL
END_METHOD

METHOD RELEASELOCK
END_METHOD

METHOD REMOVEALLELEMENTS : COLLECTION_ERROR
END_METHOD

METHOD REMOVEALLELEMENTSINTERNAL : COLLECTION_ERROR
END_METHOD

METHOD REMOVEELEMENT : COLLECTION_ERROR
VAR_INPUT
	ITFELEMENT : IElement;
END_VAR
END_METHOD

METHOD REMOVEELEMENTAT : COLLECTION_ERROR
VAR_INPUT
	UDIPOSITION : UDINT;
END_VAR
END_METHOD

METHOD REMOVEELEMENTATINTERNAL : COLLECTION_ERROR
VAR_INPUT
	UDIPOSITION : UDINT;
END_VAR
END_METHOD

METHOD SAFEELEMENTITERATOR : COLLECTION_ERROR
VAR_INPUT
	ITFITERATOR : ISafeListIterator;
END_VAR
END_METHOD

METHOD SETELEMENTAT : COLLECTION_ERROR
VAR_INPUT
	UDIPOSITION : UDINT;
	ITFELEMENT : IElement;
END_VAR
END_METHOD

METHOD SORT : COLLECTION_ERROR
END_METHOD

METHOD PRVINSTINIT : FBF.ERROR
VAR_INPUT
	ITFDATA : FBF.IData;
END_VAR
END_METHOD

(* ---- SORTEDLISTFACTORY.fb ---- *)
FUNCTION_BLOCK SORTEDLISTFACTORY EXTENDS FactoryBase
VAR
	PRVINSTCOUNT : CAA.COUNT;
	PRVINSTPOOLEXTENDSFACTOR : USINT;
	PRVINSTSIZE : CAA.SIZE;
END_VAR
END_FUNCTION_BLOCK

METHOD CREATE : ISortedList3
VAR_INPUT
	UDIMAXELEMENTS : UDINT;
END_VAR
VAR_OUTPUT
	EERROR : FBF.ERROR;
END_VAR
END_METHOD

METHOD CREATEDYNAMICLIST : ISortedList2
VAR_INPUT
	UDIINITIALSIZE : UDINT;
	UIGROWFACTOR : UINT;
END_VAR
VAR_OUTPUT
	EERROR : FBF.ERROR;
END_VAR
END_METHOD

(* ---- STACK.fb ---- *)
FUNCTION_BLOCK STACK EXTENDS InstanceBase
VAR_INPUT
	PAELEMENTS : POINTER TO IElement;
	UDIMAXELEMENTS : UDINT;
END_VAR
VAR
	_DIMAXPOSITION : DINT := -1;
	_SNAME : STRING := 'List';
	RESULT : RTS_IEC_RESULT;
	_XWPOINTERTOTHIS : __XWORD := THIS;
	_BYLOCK : BYTE;
	_ULINTCOUNTMODS : ULINT;
	_UIGROWFACTOR : UINT := 1;
	_LOCKWAITTIME : SYSTIME := Variables.g_LockWaitTime;
	COUNTMODIFICATIONS : ULINT;
	LOCKWAITTIME : SYSTIME;
END_VAR
END_FUNCTION_BLOCK

METHOD ADDELEMENT : COLLECTION_ERROR
VAR_INPUT
	ITFELEMENT : IElement;
END_VAR
END_METHOD

METHOD CONTAINSELEMENT : COLLECTION_ERROR
VAR_INPUT
	ITFELEMENT : IElement;
END_VAR
VAR_OUTPUT
	XRESULT : BOOL;
END_VAR
END_METHOD

METHOD CONTAINSVALUE : COLLECTION_ERROR
VAR_INPUT
	ITFELEMENT : IElement;
END_VAR
VAR_OUTPUT
	XRESULT : BOOL;
END_VAR
END_METHOD

METHOD COUNTELEMENTS : UDINT
END_METHOD

METHOD DISPOSE : BOOL
END_METHOD

METHOD ELEMENTCOMPARETO : INT
VAR_INPUT
	ITFELEMENT : IElement;
END_VAR
END_METHOD

METHOD ELEMENTEQUALS : BOOL
VAR_INPUT
	ITFELEMENT : IElement;
END_VAR
END_METHOD

METHOD ELEMENTHASHCODE : LINT
END_METHOD

METHOD ELEMENTITERATOR : COLLECTION_ERROR
VAR_INPUT
	ITFITERATOR : IIterator;
END_VAR
END_METHOD

METHOD LOCK : BOOL
END_METHOD

METHOD PEEK : COLLECTION_ERROR
VAR_OUTPUT
	ITFELEMENT : IElement;
END_VAR
END_METHOD

METHOD POP : COLLECTION_ERROR
VAR_OUTPUT
	ITFELEMENT : IElement;
END_VAR
END_METHOD

METHOD REALLOC : BOOL
END_METHOD

METHOD RELEASELOCK
END_METHOD

METHOD REMOVEALLELEMENTS : COLLECTION_ERROR
END_METHOD

METHOD REMOVEALLELEMENTSINTERNAL : COLLECTION_ERROR
END_METHOD

METHOD REMOVEELEMENT : COLLECTION_ERROR
VAR_INPUT
	ITFELEMENT : IElement;
END_VAR
END_METHOD

METHOD REMOVEELEMENTATINTERNAL : COLLECTION_ERROR
VAR_INPUT
	UDIPOSITION : UDINT;
END_VAR
END_METHOD

METHOD SAFEELEMENTITERATOR : COLLECTION_ERROR
VAR_INPUT
	ITFITERATOR : ISafeListIterator;
END_VAR
END_METHOD

METHOD PRVINSTINIT : FBF.ERROR
VAR_INPUT
	ITFDATA : FBF.IData;
END_VAR
END_METHOD

(* ---- STACKFACTORY.fb ---- *)
FUNCTION_BLOCK STACKFACTORY EXTENDS FactoryBase
VAR
	PRVINSTCOUNT : CAA.COUNT;
	PRVINSTPOOLEXTENDSFACTOR : USINT;
	PRVINSTSIZE : CAA.SIZE;
END_VAR
END_FUNCTION_BLOCK

METHOD CREATE : IStack3
VAR_INPUT
	UDIMAXELEMENTS : UDINT;
END_VAR
VAR_OUTPUT
	EERROR : FBF.ERROR;
END_VAR
END_METHOD

METHOD CREATEDYNAMICSTACK : IStack2
VAR_INPUT
	UDIINITIALSIZE : UDINT;
	UIGROWFACTOR : UINT;
END_VAR
VAR_OUTPUT
	EERROR : FBF.ERROR;
END_VAR
END_METHOD

(* ---- STRINGDATA.fb ---- *)
FUNCTION_BLOCK STRINGDATA EXTENDS InstanceData
VAR_INPUT
	SVALUE : STRING;
END_VAR
END_FUNCTION_BLOCK

(* ---- STRINGELEMENT.fb ---- *)
FUNCTION_BLOCK STRINGELEMENT EXTENDS InstanceBase
VAR_INPUT
	SVALUE : STRING;
END_VAR
VAR
	STRINGVALUE : STRING;
END_VAR
END_FUNCTION_BLOCK

METHOD ELEMENTCOMPARETO : INT
VAR_INPUT
	ITFELEMENT : IElement;
END_VAR
END_METHOD

METHOD ELEMENTEQUALS : BOOL
VAR_INPUT
	ITFELEMENT : IElement;
END_VAR
END_METHOD

METHOD ELEMENTHASHCODE : LINT
END_METHOD

METHOD PRVINSTINIT : FBF.ERROR
VAR_INPUT
	ITFDATA : FBF.IData;
END_VAR
END_METHOD

(* ---- STRINGELEMENTFACTORY.fb ---- *)
FUNCTION_BLOCK STRINGELEMENTFACTORY EXTENDS FactoryBase
VAR
	PRVINSTCOUNT : CAA.COUNT;
	PRVINSTPOOLEXTENDSFACTOR : USINT;
	PRVINSTSIZE : CAA.SIZE;
END_VAR
END_FUNCTION_BLOCK

METHOD CREATE : IStringElement
VAR_INPUT
	SVALUE : STRING;
END_VAR
VAR_OUTPUT
	EERROR : FBF.ERROR;
END_VAR
END_METHOD

(* ---- TIMEDATA.fb ---- *)
FUNCTION_BLOCK TIMEDATA EXTENDS InstanceData
VAR_INPUT
	TVALUE : TIME;
END_VAR
END_FUNCTION_BLOCK

(* ---- TIMEELEMENT.fb ---- *)
FUNCTION_BLOCK TIMEELEMENT EXTENDS InstanceBase
VAR_INPUT
	TVALUE : TIME;
END_VAR
VAR
	TIMEVALUE : TIME;
END_VAR
END_FUNCTION_BLOCK

METHOD ELEMENTCOMPARETO : INT
VAR_INPUT
	ITFELEMENT : IElement;
END_VAR
END_METHOD

METHOD ELEMENTEQUALS : BOOL
VAR_INPUT
	ITFELEMENT : IElement;
END_VAR
END_METHOD

METHOD ELEMENTHASHCODE : LINT
END_METHOD

METHOD PRVINSTINIT : FBF.ERROR
VAR_INPUT
	ITFDATA : FBF.IData;
END_VAR
END_METHOD

(* ---- TIMEELEMENTFACTORY.fb ---- *)
FUNCTION_BLOCK TIMEELEMENTFACTORY EXTENDS FactoryBase
VAR
	PRVINSTCOUNT : CAA.COUNT;
	PRVINSTPOOLEXTENDSFACTOR : USINT;
	PRVINSTSIZE : CAA.SIZE;
END_VAR
END_FUNCTION_BLOCK

METHOD CREATE : ITimeElement
VAR_INPUT
	TVALUE : TIME;
END_VAR
VAR_OUTPUT
	EERROR : FBF.ERROR;
END_VAR
END_METHOD

(* ---- TREENODE.fb ---- *)
FUNCTION_BLOCK TREENODE EXTENDS InstanceBase
VAR
	_LINKEDLIST : LinkedList;
	_XWPOINTERTOTHIS : __XWORD := THIS;
	_BYLOCK : BYTE;
	_ITFELEMENT : IElement;
	_ITFPARENTNODE : ITreeNode;
	_LOCKWAITTIME : SYSTIME := Variables.g_LockWaitTime;
	ELEMENT : IElement;
	LOCKWAITTIME : SYSTIME;
END_VAR
END_FUNCTION_BLOCK

METHOD ADDCHILD : COLLECTION_ERROR
VAR_INPUT
	ITFELEMENT : IElement;
END_VAR
VAR_OUTPUT
	ITFTREENODE : ITreeNode;
END_VAR
END_METHOD

METHOD CHILDREN : COLLECTION_ERROR
VAR_INPUT
	ITFITERATOR : IIterator;
END_VAR
END_METHOD

METHOD CONTAINSCHILD : COLLECTION_ERROR
VAR_INPUT
	ITFELEMENT : IElement;
END_VAR
VAR_OUTPUT
	XRESULT : BOOL;
END_VAR
END_METHOD

METHOD CONTAINSSUBNODE : COLLECTION_ERROR
VAR_INPUT
	ITFTREENODE : ITreeNode;
END_VAR
VAR_OUTPUT
	XRESULT : BOOL;
END_VAR
END_METHOD

METHOD COUNTCHILDREN : UDINT
END_METHOD

METHOD DISPOSE : BOOL
END_METHOD

METHOD ELEMENTCOMPARETO : INT
VAR_INPUT
	ITFELEMENT : IElement;
END_VAR
END_METHOD

METHOD ELEMENTEQUALS : BOOL
VAR_INPUT
	ITFELEMENT : IElement;
END_VAR
END_METHOD

METHOD ELEMENTHASHCODE : LINT
END_METHOD

METHOD LOCK : BOOL
END_METHOD

METHOD MOVENODE : COLLECTION_ERROR
VAR_INPUT
	ITFTARGETTREENODE : ITreeNode;
END_VAR
END_METHOD

METHOD PARENT : COLLECTION_ERROR
VAR_OUTPUT
	ITFPARENT : ITreeNode;
END_VAR
END_METHOD

METHOD RELEASELOCK
END_METHOD

METHOD REMOVECHILD : COLLECTION_ERROR
VAR_INPUT
	ITFELEMENT : IElement;
END_VAR
END_METHOD

METHOD ROOTNODE : COLLECTION_ERROR
VAR_OUTPUT
	ITFROOTNODE : ITreeNode;
END_VAR
END_METHOD

METHOD SAFECHILDREN : COLLECTION_ERROR
VAR_INPUT
	ITFITERATOR : ISafeLinkedListIterator;
END_VAR
END_METHOD

METHOD PRVINSTINIT : FBF.ERROR
VAR_INPUT
	ITFDATA : FBF.IData;
END_VAR
END_METHOD

(* ---- TREENODEARGS.fb ---- *)
FUNCTION_BLOCK TREENODEARGS EXTENDS InstanceData
VAR_INPUT
	ITFELEMENT : IElement;
	ITFPARENT : ITreeNode;
END_VAR
END_FUNCTION_BLOCK

(* ---- TREENODEFACTORY.fb ---- *)
FUNCTION_BLOCK TREENODEFACTORY EXTENDS FactoryBase
VAR
	PRVINSTCOUNT : CAA.COUNT;
	PRVINSTPOOLEXTENDSFACTOR : USINT;
	PRVINSTSIZE : CAA.SIZE;
END_VAR
END_FUNCTION_BLOCK

METHOD CREATE : ITreeNode2
VAR_INPUT
	ITFELEMENT : IElement;
END_VAR
VAR_OUTPUT
	EERROR : FBF.ERROR;
END_VAR
END_METHOD

METHOD CREATEINTERNAL : ITreeNode2
VAR_INPUT
	ITFELEMENT : IElement;
	ITFPARENT : ITreeNode;
END_VAR
VAR_OUTPUT
	EERROR : FBF.ERROR;
END_VAR
END_METHOD

(* ---- UDINTDATA.fb ---- *)
FUNCTION_BLOCK UDINTDATA EXTENDS InstanceData
VAR_INPUT
	UDIVALUE : UDINT;
END_VAR
END_FUNCTION_BLOCK

(* ---- UDINTELEMENT.fb ---- *)
FUNCTION_BLOCK UDINTELEMENT EXTENDS InstanceBase
VAR_INPUT
	UDIVALUE : UDINT;
END_VAR
VAR
	UDINTVALUE : UDINT;
END_VAR
END_FUNCTION_BLOCK

METHOD ELEMENTCOMPARETO : INT
VAR_INPUT
	ITFELEMENT : IElement;
END_VAR
END_METHOD

METHOD ELEMENTEQUALS : BOOL
VAR_INPUT
	ITFELEMENT : IElement;
END_VAR
END_METHOD

METHOD ELEMENTHASHCODE : LINT
END_METHOD

METHOD PRVINSTINIT : FBF.ERROR
VAR_INPUT
	ITFDATA : FBF.IData;
END_VAR
END_METHOD

(* ---- UDINTELEMENTFACTORY.fb ---- *)
FUNCTION_BLOCK UDINTELEMENTFACTORY EXTENDS FactoryBase
VAR
	PRVINSTCOUNT : CAA.COUNT;
	PRVINSTPOOLEXTENDSFACTOR : USINT;
	PRVINSTSIZE : CAA.SIZE;
END_VAR
END_FUNCTION_BLOCK

METHOD CREATE : IUdintElement
VAR_INPUT
	UDIVALUE : UDINT;
END_VAR
VAR_OUTPUT
	EERROR : FBF.ERROR;
END_VAR
END_METHOD

(* ---- UINTDATA.fb ---- *)
FUNCTION_BLOCK UINTDATA EXTENDS InstanceData
VAR_INPUT
	UIVALUE : UINT;
END_VAR
END_FUNCTION_BLOCK

(* ---- UINTELEMENT.fb ---- *)
FUNCTION_BLOCK UINTELEMENT EXTENDS InstanceBase
VAR_INPUT
	UIVALUE : UINT;
END_VAR
VAR
	UINTVALUE : UINT;
END_VAR
END_FUNCTION_BLOCK

METHOD ELEMENTCOMPARETO : INT
VAR_INPUT
	ITFELEMENT : IElement;
END_VAR
END_METHOD

METHOD ELEMENTEQUALS : BOOL
VAR_INPUT
	ITFELEMENT : IElement;
END_VAR
END_METHOD

METHOD ELEMENTHASHCODE : LINT
END_METHOD

METHOD PRVINSTINIT : FBF.ERROR
VAR_INPUT
	ITFDATA : FBF.IData;
END_VAR
END_METHOD

(* ---- UINTELEMENTFACTORY.fb ---- *)
FUNCTION_BLOCK UINTELEMENTFACTORY EXTENDS FactoryBase
VAR
	PRVINSTCOUNT : CAA.COUNT;
	PRVINSTPOOLEXTENDSFACTOR : USINT;
	PRVINSTSIZE : CAA.SIZE;
END_VAR
END_FUNCTION_BLOCK

METHOD CREATE : IUintElement
VAR_INPUT
	UIVALUE : UINT;
END_VAR
VAR_OUTPUT
	EERROR : FBF.ERROR;
END_VAR
END_METHOD

(* ---- ULINTDATA.fb ---- *)
FUNCTION_BLOCK ULINTDATA EXTENDS InstanceData
VAR_INPUT
	ULIVALUE : ULINT;
END_VAR
END_FUNCTION_BLOCK

(* ---- ULINTELEMENT.fb ---- *)
FUNCTION_BLOCK ULINTELEMENT EXTENDS InstanceBase
VAR_INPUT
	ULIVALUE : ULINT;
END_VAR
VAR
	ULINTVALUE : ULINT;
END_VAR
END_FUNCTION_BLOCK

METHOD ELEMENTCOMPARETO : INT
VAR_INPUT
	ITFELEMENT : IElement;
END_VAR
END_METHOD

METHOD ELEMENTEQUALS : BOOL
VAR_INPUT
	ITFELEMENT : IElement;
END_VAR
END_METHOD

METHOD ELEMENTHASHCODE : LINT
END_METHOD

METHOD PRVINSTINIT : FBF.ERROR
VAR_INPUT
	ITFDATA : FBF.IData;
END_VAR
END_METHOD

(* ---- ULINTELEMENTFACTORY.fb ---- *)
FUNCTION_BLOCK ULINTELEMENTFACTORY EXTENDS FactoryBase
VAR
	PRVINSTCOUNT : CAA.COUNT;
	PRVINSTPOOLEXTENDSFACTOR : USINT;
	PRVINSTSIZE : CAA.SIZE;
END_VAR
END_FUNCTION_BLOCK

METHOD CREATE : IUlintElement
VAR_INPUT
	ULIVALUE : ULINT;
END_VAR
VAR_OUTPUT
	EERROR : FBF.ERROR;
END_VAR
END_METHOD

(* ---- WSTRINGDATA.fb ---- *)
FUNCTION_BLOCK WSTRINGDATA EXTENDS InstanceData
VAR_INPUT
	WSVALUE : WSTRING;
END_VAR
END_FUNCTION_BLOCK

(* ---- WSTRINGELEMENT.fb ---- *)
FUNCTION_BLOCK WSTRINGELEMENT EXTENDS InstanceBase
VAR_INPUT
	WSVALUE : WSTRING;
END_VAR
VAR
	WSTRINGVALUE : WSTRING;
END_VAR
END_FUNCTION_BLOCK

METHOD ELEMENTCOMPARETO : INT
VAR_INPUT
	ITFELEMENT : IElement;
END_VAR
END_METHOD

METHOD ELEMENTEQUALS : BOOL
VAR_INPUT
	ITFELEMENT : IElement;
END_VAR
END_METHOD

METHOD ELEMENTHASHCODE : LINT
END_METHOD

METHOD PRVINSTINIT : FBF.ERROR
VAR_INPUT
	ITFDATA : FBF.IData;
END_VAR
END_METHOD

(* ---- WSTRINGELEMENTFACTORY.fb ---- *)
FUNCTION_BLOCK WSTRINGELEMENTFACTORY EXTENDS FactoryBase
VAR
	PRVINSTCOUNT : CAA.COUNT;
	PRVINSTPOOLEXTENDSFACTOR : USINT;
	PRVINSTSIZE : CAA.SIZE;
END_VAR
END_FUNCTION_BLOCK

METHOD CREATE : IWStringElement
VAR_INPUT
	WSVALUE : WSTRING;
END_VAR
VAR_OUTPUT
	EERROR : FBF.ERROR;
END_VAR
END_METHOD
